FUNCTION_BLOCK EP_Pump (* The equipment as its skills see it, the same in every skill that uses it: plays a command (its output values, phase by phase) on the equipment's command channel, and gives the equipment's newest state. Technical: Pump as its skills see it: a command on the socket Skill (AEquipment: SEND, PLAYED when all phases are out) goes out on its command channel; STATE gives its inputs and holder *)
  (* Standard: 61499-2 *)
  (* Version 0.1, 2026-09-28, Project contributors, AAU Smart Production Lab *)
  PACKAGE filling;
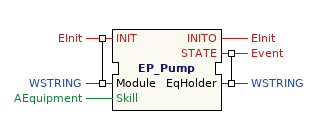
  EVENT_INPUT
    INIT : EInit WITH Module; (* Initialise: name the equipment's channels and listen to its state *)
  END_EVENT
  EVENT_OUTPUT
    INITO : EInit; (* Initialised: the next block of the INIT chain goes on *)
    STATE WITH EqHolder; (* The equipment's newest state: its inputs and who holds it *)
  END_EVENT
  VAR_INPUT
    Module : WSTRING; (* The module's name; its local channels are named after it (loc[<Module>/...]) *)
  END_VAR
  VAR_OUTPUT
    EqHolder : WSTRING; (* Who holds the equipment now (empty: free) *)
  END_VAR
  SOCKETS
    Skill : modlib::AEquipment; (* From a skill's run (AEquipment): the commands to play, PLAYED back *)
  END_SOCKETS
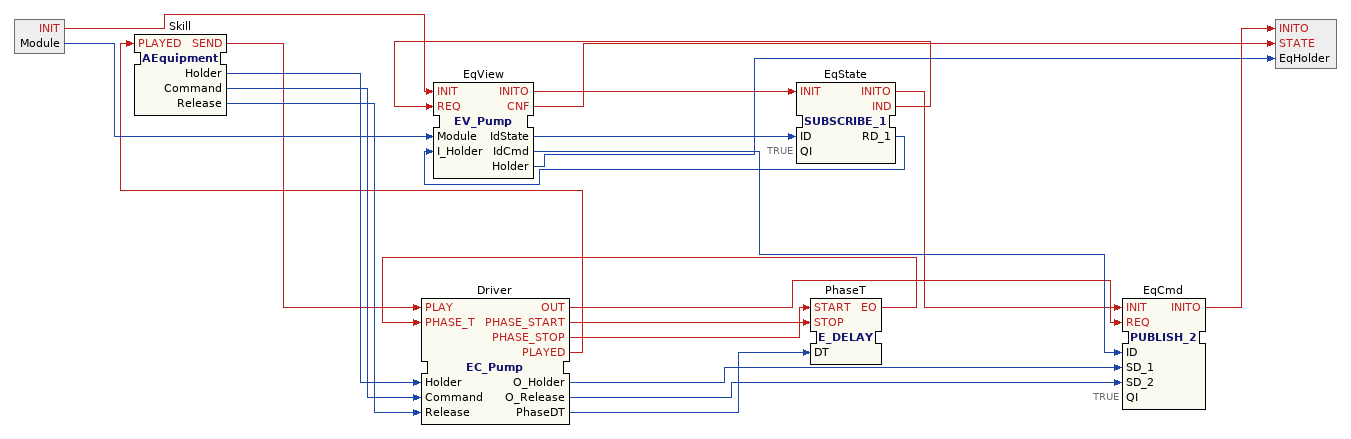
  (* Group StateIn: The equipment's state in: its inputs and who holds it, from its state channel *)
  (* Group CommandOut: A command out: its output values, phase by phase (the command table), on the command channel *)
  FBS
    EqView : filling::EV_Pump; (* Names the equipment's channels, and unpacks its state into named values. *) {SET_ATTRIBUTE(GroupName, StateIn)}
    EqState : iec61499::net::SUBSCRIBE_1(QI := TRUE); (* Listens to the equipment's state channel: its inputs and who holds it. *) {SET_ATTRIBUTE(GroupName, StateIn)}
    Driver : filling::EC_Pump; (* The equipment's command table (EC_): turns a command into output values, phase by phase. *) {SET_ATTRIBUTE(GroupName, CommandOut)}
    PhaseT : iec61499::events::E_DELAY; (* Times the phases of a command. *) {SET_ATTRIBUTE(GroupName, CommandOut)}
    EqCmd : iec61499::net::PUBLISH_2(QI := TRUE); (* Sends the output values and the holder's name to the equipment block on its command channel. *) {SET_ATTRIBUTE(GroupName, CommandOut)}
  END_FBS
  EVENT_CONNECTIONS
    INIT TO EqView.INIT;
    EqView.INITO TO EqState.INIT;
    EqState.INITO TO EqCmd.INIT;
    EqCmd.INITO TO INITO;
    EqState.IND TO EqView.REQ;
    EqView.CNF TO STATE;
    Skill.SEND TO Driver.PLAY;
    Driver.OUT TO EqCmd.REQ;
    Driver.PHASE_START TO PhaseT.START;
    Driver.PHASE_STOP TO PhaseT.STOP;
    PhaseT.EO TO Driver.PHASE_T;
    Driver.PLAYED TO Skill.PLAYED;
  END_CONNECTIONS
  DATA_CONNECTIONS
    Module TO EqView.Module;
    EqView.IdState TO EqState.ID;
    EqView.IdCmd TO EqCmd.ID;
    EqState.RD_1 TO EqView.I_Holder;
    EqView.Holder TO EqHolder;
    Skill.Holder TO Driver.Holder;
    Skill.Command TO Driver.Command;
    Skill.Release TO Driver.Release;
    Driver.O_Holder TO EqCmd.SD_1;
    Driver.O_Release TO EqCmd.SD_2;
    Driver.PhaseDT TO PhaseT.DT;
  END_CONNECTIONS
END_FUNCTION_BLOCK
